(* IEC 61131-3 sources: JingjiangMoonbox/Application/Application/任务列表/TensionTask/电机运动/SetMode, 4 files *)

(* ---- SetPrfGantryTrapModePrm.st ---- *)
(*@CES
Name=SetPrfGantryTrapModePrm
Type=FunctionBlock
TypeGuid=6f9dac99-8de1-4efc-8465-68ac443b7d08
Guid=46cb849a-922f-49f0-be65-4966a012b8cb
HasDeclaration=True
HasImplementation=True
*)
{DECLARATION}
FUNCTION SetPrfGantryTrapModePrm : INT
VAR_INPUT
	i_iCoreId:INT;							//前64轴核号为1，后64轴轴号为2
	i_iGroupId : INT;
	i_iAxisMaster:INT;
	i_iAxisSlaver:INT;
	i_iAxisMasterVirtual:INT;//主轴叠加轴轴号；
	i_diSyncErrorLimit : DINT;
END_VAR
VAR
	iRtn:INT:=0;
	STGantryPrmPro : TGantryPrmPro;
	STPidAlign : TPidAlign;
END_VAR

{IMPLEMENTATION}
// SysMemSet(ADR(STGantryPrmPro),0,SIZEOF(STGantryPrmPro));
//
// STGantryPrmPro.mode := GANTRY_MODE_NONE;									//龙门模式  20开环龙门模式  勿改
// STGantryPrmPro.master :=i_iAxisMaster;						//主轴轴号
// STGantryPrmPro.slave := i_iAxisSlaver;							//从轴轴号
// STGantryPrmPro.reserve[0] := i_iAxisMasterVirtual;				//主轴叠加轴轴号；此数组从0开始，一定要注意
// STGantryPrmPro.reserve[1] := 0;								//必须为0
// STGantryPrmPro.reserve[2] := 0;								//必须为0
// STGantryPrmPro.syncErrorLimit := i_diSyncErrorLimit;					//龙门最大差值
//
// STGantryPrmPro.gantryMasterPid.kp := 1;
// STGantryPrmPro.gantrySlavePid.kp := 1;
// STGantryPrmPro.masterPid.kp := 1;
// STGantryPrmPro.slavePid.kp := 1;
// iRtn := GTN_SetGantryPrmPro(core:= i_iCoreId, group:=i_iGroupId, pGantryPrmPro:= ADR(STGantryPrmPro)) + iRtn;

SysMemSet(ADR(STGantryPrmPro),0,SIZEOF(STGantryPrmPro));

STGantryPrmPro.mode := 20;									//龙门模式  20开环龙门模式  勿改
STGantryPrmPro.master :=i_iAxisMaster;						//主轴轴号
STGantryPrmPro.slave := i_iAxisSlaver;							//从轴轴号
STGantryPrmPro.reserve[0] := i_iAxisMasterVirtual;				//主轴叠加轴轴号；此数组从0开始，一定要注意
STGantryPrmPro.reserve[1] := 0;								//必须为0
STGantryPrmPro.reserve[2] := 0;								//必须为0
STGantryPrmPro.syncErrorLimit := i_diSyncErrorLimit;					//龙门最大差值

STGantryPrmPro.gantryMasterPid.kp := 1;
STGantryPrmPro.gantrySlavePid.kp := 1;
STGantryPrmPro.masterPid.kp := 1;
STGantryPrmPro.slavePid.kp := 1;
//
// STPidAlign.kp := 1;
// STPidAlign.ki := 1;
// STPidAlign.kd := 1;
// STPidAlign.kaff := 1;
// STPidAlign.kvff := 1;
// STPidAlign.derivativeLimit := 1;
// STPidAlign.integralLimit := 1;
// STPidAlign.s_limit := 1;
// STPidAlign.reserve[1] := 0;
// STPidAlign.reserve[2] := 0;

// SysMemCpy(ADR(STGantryPrmPro.gantryMasterPid),ADR(STPidAlign),SIZEOF(STPidAlign));
// SysMemCpy(ADR(STGantryPrmPro.gantrySlavePid),ADR(STPidAlign),SIZEOF(STPidAlign));
// SysMemCpy(ADR(STGantryPrmPro.masterPid),ADR(STPidAlign),SIZEOF(STPidAlign));
// SysMemCpy(ADR(STGantryPrmPro.slavePid),ADR(STPidAlign),SIZEOF(STPidAlign));

iRtn := GTN_SetGantryPrmPro(core:= i_iCoreId, group:=i_iGroupId, pGantryPrmPro:= ADR(STGantryPrmPro)) + iRtn;

iRtn := SetPrfTrapModePrm(
				i_iCoreId:= i_iCoreId,
				i_iAxisId:= i_iAxisMaster,
				i_lrVel:= 100,//i_pastTStTrapParamUser^[iCnt_TrapAxis].lrVel,
				i_lrAcc:= 1,//i_pastTStTrapParamUser^[iCnt_TrapAxis].lrAcc,
				i_lrDec:= 1,//i_pastTStTrapParamUser^[iCnt_TrapAxis].lrDec,
				i_iSmoothTime:= 0) + iRtn;//i_pastTStTrapParamUser^[iCnt_TrapAxis].iSmoothTime);

iRtn := SetPrfTrapModePrm(
				i_iCoreId:= i_iCoreId,
				i_iAxisId:= i_iAxisSlaver,
				i_lrVel:= 100,//i_pastTStTrapParamUser^[iCnt_TrapAxis].lrVel,
				i_lrAcc:= 1,//i_pastTStTrapParamUser^[iCnt_TrapAxis].lrAcc,
				i_lrDec:= 1,//i_pastTStTrapParamUser^[iCnt_TrapAxis].lrDec,
				i_iSmoothTime:= 0) + iRtn;//i_pastTStTrapParamUser^[iCnt_TrapAxis].iSmoothTime);

iRtn := SetPrfTrapModePrm(
				i_iCoreId:= i_iCoreId,
				i_iAxisId:= i_iAxisMasterVirtual,
				i_lrVel:= 100,//i_pastTStTrapParamUser^[iCnt_TrapAxis].lrVel,
				i_lrAcc:= 1,//i_pastTStTrapParamUser^[iCnt_TrapAxis].lrAcc,
				i_lrDec:= 1,//i_pastTStTrapParamUser^[iCnt_TrapAxis].lrDec,
				i_iSmoothTime:= 0) + iRtn;//i_pastTStTrapParamUser^[iCnt_TrapAxis].iSmoothTime);

SetPrfGantryTrapModePrm:=iRtn;

(* ---- SetPrfGearModePrm.st ---- *)
(*@CES
Name=SetPrfGearModePrm
Type=FunctionBlock
TypeGuid=6f9dac99-8de1-4efc-8465-68ac443b7d08
Guid=f035424c-4733-45cb-8bf8-2e7099a0fe7e
HasDeclaration=True
HasImplementation=True
*)
{DECLARATION}
FUNCTION SetPrfGearModePrm : INT
VAR_INPUT
	i_iCore:INT;					//前64轴核号为1，后64轴轴号为2
	i_iAxisId:INT;
	i_iMasterIndex:INT;		//主轴索引
	i_diMasterEven:DINT;	//主轴转数
	i_diSlaveEven:DINT;		//从轴转数
	i_diMasterSlope:DINT;	//离合区
	i_xMasterType : BOOL;
END_VAR
VAR
	iRtn: INT;
	iMasterType : INT;
END_VAR

{IMPLEMENTATION}
iRtn :=  GTN_PrfGear(i_iCore,i_iAxisId,0) + iRtn;
// 设置电子齿轮运动参数
IF i_xMasterType THEN
	iMasterType := GEAR_MASTER_AXIS;
ELSE
	iMasterType := GEAR_MASTER_AXIS_OTHER;
END_IF
iMasterType := GEAR_MASTER_AXIS;
iRtn :=  GTN_SetGearMaster(
		core:= i_iCore,
		profile:= i_iAxisId,
		masterIndex:= i_iMasterIndex,
		masterType:= iMasterType,
		masterItem:= 0) + iRtn;

iRtn :=  GTN_SetGearRatio(
		core:= i_iCore,
		profile:= i_iAxisId,
		masterEven:= i_diMasterEven, 					//主轴转数
		slaveEven:= i_diSlaveEven, 						//对应从轴转数
		masterSlope:= i_diMasterSlope) + iRtn;

SetPrfGearModePrm:=iRtn;

(* ---- SetPrfJogModePrm.st ---- *)
(*@CES
Name=SetPrfJogModePrm
Type=FunctionBlock
TypeGuid=6f9dac99-8de1-4efc-8465-68ac443b7d08
Guid=a1a4e312-954b-4b17-a8ec-a6ba64bc8c04
HasDeclaration=True
HasImplementation=True
*)
{DECLARATION}
FUNCTION SetPrfJogModePrm : INT
VAR_INPUT
	i_iCore:INT;							//前64轴核号为1，后64轴轴号为2
	i_iAxisId:INT;
	i_lrAcc:LREAL;
	i_lrDec:LREAL;
	i_rSmooth: REAL;
END_VAR
VAR
	iRtn:INT;
	stJogPrm:TJogPrm;
END_VAR

{IMPLEMENTATION}
iRtn :=  GTN_PrfJog(i_iCore,i_iAxisId) + iRtn;

// 读取点位运动参数(需要读取所有运动参数到上位机变量)
iRtn :=  GTN_GetJogPrm(i_iCore,i_iAxisId, ADR(stJogPrm)) + iRtn;

// 设置需要修改的运动参数
stJogPrm.acc := i_lrAcc;
stJogPrm.dec := i_lrDec;
stJogPrm.smooth := i_rSmooth;

// 设置点位运动参数
iRtn :=  GTN_SetJogPrm(i_iCore,i_iAxisId,ADR(stJogPrm)) + iRtn;

SetPrfJogModePrm:=iRtn;

(* ---- SetPrfTrapModePrm.st ---- *)
(*@CES
Name=SetPrfTrapModePrm
Type=FunctionBlock
TypeGuid=6f9dac99-8de1-4efc-8465-68ac443b7d08
Guid=a2a95545-544a-475f-b543-56a661f67a2d
HasDeclaration=True
HasImplementation=True
*)
{DECLARATION}
FUNCTION SetPrfTrapModePrm : INT
VAR_INPUT
	i_iCoreId:INT;						//前64轴核号为1，后64轴轴号为2
	i_iAxisId:INT;
	i_lrVel:LREAL;
	i_lrAcc:LREAL;
	i_lrDec:LREAL;
	i_iSmoothTime: INT;
	//i_paiRtn : POINTER TO ARRAY [1..10] OF INT;
END_VAR
VAR
	iN : INT;
	aiRtn : ARRAY [1..10] OF INT;
	stTrapPrm : TTrapPrm;
END_VAR

{IMPLEMENTATION}
aiRtn[1] :=  GTN_PrfTrap(i_iCoreId,i_iAxisId);

// 读取点位运动参数(需要读取所有运动参数到上位机变量)
aiRtn[2] :=  GTN_GetTrapPrm(i_iCoreId,i_iAxisId, ADR(stTrapPrm));

// 设置需要修改的运动参数
stTrapPrm.acc := i_lrAcc;
stTrapPrm.dec := i_lrDec;
stTrapPrm.velStart := 0;
stTrapPrm.smoothTime := i_iSmoothTime;

// 设置点位运动参数
aiRtn[3] :=  GTN_SetTrapPrm(i_iCoreId,i_iAxisId,ADR(stTrapPrm));

aiRtn[4] := GTN_SetVel(i_iCoreId,i_iAxisId,i_lrVel);

SetPrfTrapModePrm:=aiRtn[1]+aiRtn[2]+aiRtn[3]+aiRtn[4];

// FOR iN := 1 TO 10 BY 1 DO
// 	i_paiRtn^[iN] := aiRtn[iN];
// END_FOR
